Fanuc KAREL source: KA00184.KL

PROGRAM KA00184
%NOLOCKGROUP
VAR
  SRC: ARRAY[4] OF BYTE
  DST: ARRAY[4] OF STRING[20]
BEGIN
  DST = SRC
END KA00184
